Staubli VAL3: utImage.dtx

public utAppearance Appearance
  [0]
    string sBackgroundColour
    bool bVisibility
public utBorder Border
  [0]
    string sBorderColour
    string sBorderStyle
    num nBorderWidth
public utCommon Common
  [0]
    string sSourceImage
    string sID
    string sClass
    string sPage
public utEvents Events
  [0]
    bool bClick
    bool bMouseDown
    bool bMouseUp
public utData Data
  [0]
    num nVal
    bool bStatus
    string sSourceImg1
    string sSourceImg2
